FUNCTION_BLOCK Controle_Gradeamento (* Comandos do gradeamento mecanizado (padrao Grade_Comandos do legado): ciclo remoto e setpoints de diferencial de nivel das grades *)
  (* Standard: 61499-2 *)
  (* Version 1.0, 21/10/2026, Hidryco, Hidryco, 1.0: Comandos do gradeamento mecanizado (padrao Grade_Comandos do legado): ciclo remoto e setpoints de diferencial de nivel das grades *)
  PACKAGE Hidryco.HidrycoLib;
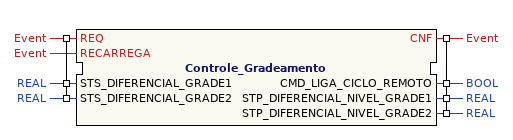
  EVENT_INPUT
    REQ WITH STS_DIFERENCIAL_GRADE1, STS_DIFERENCIAL_GRADE2; (* Status vindo do processo *)
    RECARREGA; (* Reenvia os ajustes persistentes (chamado no fim do INIT do processo) *)
  END_EVENT
  EVENT_OUTPUT
    CNF WITH CMD_LIGA_CICLO_REMOTO, STP_DIFERENCIAL_NIVEL_GRADE1, STP_DIFERENCIAL_NIVEL_GRADE2; (* Ajustes para o processo (mudanca na IHM, OPC UA ou recarga) *)
  END_EVENT
  VAR_INPUT
    STS_DIFERENCIAL_GRADE1 : REAL; (* Nivel diferencial da grade 1 agora (%) *)
    STS_DIFERENCIAL_GRADE2 : REAL; (* Nivel diferencial da grade 2 agora (%) *)
  END_VAR
  VAR_OUTPUT
    CMD_LIGA_CICLO_REMOTO : BOOL; (* Ciclo remoto *)
    STP_DIFERENCIAL_NIVEL_GRADE1 : REAL; (* Diferencial de nível para limpar a grade 1 *)
    STP_DIFERENCIAL_NIVEL_GRADE2 : REAL; (* Diferencial de nível para limpar a grade 2 *)
  END_VAR
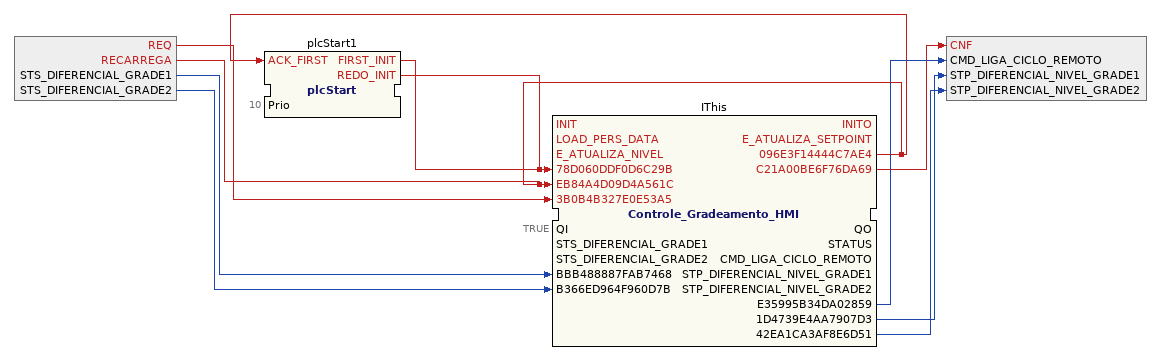
  FBS
    IThis : Controle_Gradeamento_HMI(QI := TRUE);
    plcStart1 : plcStart(Prio := 10);
  END_FBS
  EVENT_CONNECTIONS
    plcStart1.FIRST_INIT TO IThis.78D060DDF0D6C29B;
    plcStart1.REDO_INIT TO IThis.78D060DDF0D6C29B;
    IThis.096E3F14444C7AE4 TO IThis.EB84A4D09D4A561C;
    IThis.096E3F14444C7AE4 TO plcStart1.ACK_FIRST;
    RECARREGA TO IThis.EB84A4D09D4A561C;
    IThis.C21A00BE6F76DA69 TO CNF;
    REQ TO IThis.3B0B4B327E0E53A5;
  END_CONNECTIONS
  DATA_CONNECTIONS
    IThis.E35995B34DA02859 TO CMD_LIGA_CICLO_REMOTO;
    IThis.1D4739E4AA7907D3 TO STP_DIFERENCIAL_NIVEL_GRADE1;
    IThis.42EA1CA3AF8E6D51 TO STP_DIFERENCIAL_NIVEL_GRADE2;
    STS_DIFERENCIAL_GRADE1 TO IThis.BBB488887FAB7468;
    STS_DIFERENCIAL_GRADE2 TO IThis.B366ED964F960D7B;
  END_CONNECTIONS
END_FUNCTION_BLOCK
